FUNCTION FC 1 : VOID
BEGIN
NETWORK
      L I 0.0
END_FUNCTION
